Fanuc KAREL source: kx00033.KL

-- PROVISIONAL review KL for V770-1; original PC SHA256 e1684a8bb50990811f67cd31d24abe83cb7565f553f80554dcaceddecfe9d3dc
-- Incomplete behavior may be omitted. Consult companion uncertainty JSON. Do not deploy.
PROGRAM KX00033
%NOLOCKGROUP
-- UNRESOLVED_DECL I type=fa0010
-- UNRESOLVED_DECL J type=fa0010
-- UNRESOLVED_DECL B type=fa0012
-- UNRESOLVED_DECL F type=fa001d
-- UNRESOLVED_DECL S type=fa1f50
-- UNRESOLVED_DECL P type=fa0102
BEGIN
  -- UNRESOLVED_PC offsets 5-12; opcodes 9D,23
  -- UNRESOLVED_PC offsets 17-21; opcodes 7F
END KX00033
